(* IEC 61131-3 sources: Jacob-Formschaumtechnik-ISEL-CNC-Retrofit/twincat/PLC/src/6_Interfaces, 18 files *)

(* ---- E_AlarmId.st ---- *)
{attribute 'qualified_only'}
{attribute 'strict'}
TYPE E_AlarmId :
(
    None              := 0,
    SafetyOpen        := 100,  (* Sicherheitskreis offen / NOT-HALT *)
    DoorOpen          := 101,
    AirPressureLow    := 110,
    ExtractionFault   := 120,
    SpindleFuFault    := 200,
    SpindlePtcTrip    := 201,
    SpindleNoFeedback := 202,
    SpindleLockedSetup:= 203,
    AxisDriveFault    := 300,
    AxisFollowingErr  := 301,
    HwLimitHit        := 302,
    FieldbusLost      := 310,
    HomingLost        := 320,
    HmiLinkLost       := 330,
    ParamMismatch     := 900   (* Maschinen-ID oder Version passt nicht *)
) INT;
END_TYPE

(* ---- E_AlarmSlot.st ---- *)
{attribute 'qualified_only'}
{attribute 'strict'}
(* Meldekatalog: Slot-Nummer = Index in aCond von FB_AlarmList.
   Klassen siehe E_FaultClass. Texte und Abhilfe stehen in docs/Meldeliste.md (HMI-Thread). *)
TYPE E_AlarmSlot :
(
    SafetyOpen := 0,
    DoorOpen := 1,
    AirPressureLow := 2,
    ExtractionFault := 3,
    SpindleFuFault := 4,
    SpindlePtcTrip := 5,
    SpindleNoFeedback := 6,
    SpindleLockedSetup := 7,
    AxisDriveFault := 8,
    AxisFollowingErr := 9,
    HwLimitHit := 10,
    FieldbusLost := 11,
    HomingLost := 12,
    HmiLinkLost := 13,
    ParamMismatch := 14
) INT;
END_TYPE

(* ---- E_DriveVariant.st ---- *)
{attribute 'qualified_only'}
{attribute 'strict'}
(* Generische Achsschnittstelle. Variante A: CANopen DS402 ueber EL6751 (Interpolated Position
   unbestaetigt), Variante B: +-10 V Analog + Encoder-Klemmen (Rueckfall). *)
TYPE E_DriveVariant :
(
    CanopenDs402 := 0,
    AnalogEncoder := 1,
    Simulation := 2
) INT;
END_TYPE

(* ---- E_FaultClass.st ---- *)
{attribute 'qualified_only'}
{attribute 'strict'}
(* Fehlerreaktionsklassen, siehe docs/Architektur_Sicherheit.md *)
TYPE E_FaultClass :
(
    R0_Info     := 0,  (* nur anzeigen *)
    R1_Warning  := 1,  (* anzeigen, Betrieb laeuft weiter *)
    R2_FeedHold := 2,  (* gefuehrter Vorschubhalt, fortsetzbar *)
    R3_Abort    := 3,  (* gefuehrter Halt, Spindel aus, Programm beendet *)
    R4_DrivesOff := 4  (* Reglerfreigabe weg, Referenz verloren *)
) INT;
END_TYPE

(* ---- E_HomeState.st ---- *)
{attribute 'qualified_only'}
{attribute 'strict'}
TYPE E_HomeState :
(
    Open := 0,
    Running := 1,
    Done := 2,
    Error := 3
) INT;
END_TYPE

(* ---- E_MachState.st ---- *)
{attribute 'qualified_only'}
{attribute 'strict'}
TYPE E_MachState :
(
    Stopped     := 0,  (* Antriebe aus, kein Fehler *)
    Idle        := 1,  (* Antriebe bereit, kein Programm *)
    Execute     := 2,  (* Programm laeuft *)
    Held        := 3,  (* Vorschubhalt, Programm fortsetzbar *)
    Aborted     := 4,  (* Programm abgebrochen, Reset noetig *)
    EStop       := 5,  (* Sicherheitskreis offen *)
    Fault       := 6   (* Fehler R3/R4 aktiv, Quittierung noetig *)
) INT;
END_TYPE

(* ---- E_OpMode.st ---- *)
{attribute 'qualified_only'}
{attribute 'strict'}
TYPE E_OpMode :
(
    Hand  := 0,   (* Tippen, Handrad, Referenzieren *)
    Auto  := 1,   (* Programmbetrieb *)
    Setup := 2    (* Einrichten/Test: Spindel gesperrt, Einzelsatz moeglich *)
) INT;
END_TYPE

(* ---- ST_Alarm.st ---- *)
(* Eine Meldung aus der Meldeliste, Index = E_AlarmSlot *)
TYPE ST_Alarm :
STRUCT
    nId     : INT;
    eClass  : E_FaultClass;
    bActive : BOOL;          (* Ursache besteht *)
    bLatched: BOOL;          (* R3/R4 gespeichert, wartet auf Quittierung *)
END_STRUCT
END_TYPE

(* ---- ST_AxisMirror.st ---- *)
(* CNC-Spiegel fuer die HMI, Achsnummern der HMI: 1 = X (Quer), 2 = Y (Portal, Gantry), 3 = Z. *)
TYPE ST_AxisMirror :
STRUCT
    rActPosMach : LREAL;    (* mm, Maschinenkoordinate *)
    rActPosWork : LREAL;    (* mm, Werkstueckkoordinate *)
    bHomed      : BOOL;
END_STRUCT
END_TYPE

(* ---- ST_HmiCmd.st ---- *)
(* HMI -> SPS. Die HMI fordert nur an. Alle Verriegelungen liegen in der SPS. *)
TYPE ST_HmiCmd :
STRUCT
    nHeartbeat      : UINT;    (* Lebenszeichen, wird von der HMI hochgezaehlt *)
    eModeRequest    : E_OpMode;
    bStart          : BOOL;    (* Impuls *)
    bHold           : BOOL;    (* Impuls, Vorschubhalt *)
    bAbort          : BOOL;    (* Impuls *)
    bAck            : BOOL;    (* Impuls, Meldungen quittieren, Wiederanlauf *)
    bJogPlus        : BOOL;    (* gehalten, nur mit Heartbeat *)
    bJogMinus       : BOOL;
    nJogAxis        : USINT;   (* 1=X, 2=Y, 3=Z *)
    bJogRapid       : BOOL;
    bSpindleOn      : BOOL;    (* nur Hand *)
    bSpindleCcw     : BOOL;
    rSpindleSetRpm  : REAL;    (* 1/min *)
    bExtraction     : BOOL;
    bBlowAir        : BOOL;
    bVacuum         : BOOL;
    bHomeRequest    : BOOL;    (* Impuls *)
    bToolChangeDone : BOOL;    (* Impuls, Quittung manueller Werkzeugwechsel *)
    rJogStepMm      : REAL;    (* 0 = kontinuierlich, sonst 0.01 / 0.1 / 1 / 10 mm *)
    bHandwheelEnable: BOOL;    (* nur M1 mit Bestandsgeraet, [offen] *)
    nHandwheelAxis  : USINT;   (* 1=X, 2=Y, 3=Z *)
    nHandwheelRatio : USINT;   (* 1, 10, 100 *)
    bHomeAxis       : ARRAY[1..3] OF BOOL;   (* Impuls: einzelne Achse referenzieren *)
    bHomeAbort      : BOOL;    (* Impuls *)
    bSingleBlock    : BOOL;    (* Einzelsatz *)
    bDryRun         : BOOL;    (* Trockenlauf: Spindel gesperrt *)
    bOptStop        : BOOL;    (* optionaler Halt M1 *)
END_STRUCT
END_TYPE

(* ---- ST_HmiCncCmd.st ---- *)
(* HMI -> SPS *)
TYPE ST_HmiCncCmd :
STRUCT
    nOvrFeed       : UINT := 100;                (* % 0..120 *)
    nOvrRapid      : UINT := 100;                (* % 0..100 *)
    nOvrSpindle    : UINT := 100;                (* % 50..120 *)
    sProgramSelect : STRING(255);
    bProgramLoad   : BOOL;                       (* Impuls, nur im Stillstand *)
    aTool          : ARRAY[1..32] OF ST_Tool;    (* Schreibpuffer *)
    aWcs           : ARRAY[54..59] OF ST_Wcs;
    bTableWrite    : BOOL;                       (* Impuls: Puffer uebernehmen *)
    bWcsSetCurrent : BOOL;                       (* Impuls: aktuelle Position als Nullpunkt von nActWcs *)
    bWcsTableWrite : BOOL;                       (* Impuls: nur die Nullpunkte (G54..G59) aus aWcs uebernehmen. bTableWrite uebernimmt nur noch Werkzeuge (G-16) *)
    nSpeedLimitPct : UINT := 25;                 (* % 1..100, Inbetriebnahme-Begrenzung (Service). Wirkt nur nach unten auf Vorschub-/Eilgang-Override und Tippen. Anheben nur im Stillstand. *)
END_STRUCT
END_TYPE

(* ---- ST_HmiCncSts.st ---- *)
(* SPS -> HMI *)
TYPE ST_HmiCncSts :
STRUCT
    aAxis         : ARRAY[1..3] OF ST_AxisMirror;
    rGantryDiffMm : LREAL;                       (* Y1 minus Y2 *)
    nOvrFeed      : UINT;                        (* % *)
    nOvrRapid     : UINT;
    nOvrSpindle   : UINT;
    sProgramName  : STRING(80);
    nActBlock     : UDINT;
    nTotalBlocks  : UDINT;
    sBlockText    : ARRAY[0..6] OF STRING(80);   (* Index 3 = aktueller Satz *)
    rRestMm       : LREAL;
    rFeedAct      : LREAL;                       (* mm/min *)
    nActTool      : UINT;
    nActWcs       : UINT := 54;                  (* 54..59 *)
    aTool         : ARRAY[1..32] OF ST_Tool;
    aWcs          : ARRAY[54..59] OF ST_Wcs;
    bProgramLoaded: BOOL;
    bTableWriteOk : BOOL;                        (* Rueckmeldung letzter Schreibvorgang *)
    bTableWriteRejected : BOOL;                  (* abgelehnt, z. B. Programm laeuft *)
    nSpeedLimitActivePct : UINT := 25;           (* wirksame Inbetriebnahme-Begrenzung in %, nOvrFeed/nOvrRapid sind bereits damit begrenzt *)
END_STRUCT
END_TYPE

(* ---- ST_HmiJournal.st ---- *)
(* Meldejournal fuer die HMI (Befund 21, LH-2.9.2). Ringpuffer der letzten 100 kommenden Meldungen.
   nHead zeigt auf den naechsten freien Platz, der juengste Eintrag steht bei (nHead + 99) MOD 100.
   nSeq zaehlt jeden neuen Eintrag hoch, die HMI liest nur bei Aenderung. *)
TYPE ST_HmiJournal :
STRUCT
    aEntry   : ARRAY[0..99] OF ST_JournalEntry;
    nHead    : UINT;
    nEntries : UINT;
    nSeq     : UDINT;
END_STRUCT
END_TYPE

(* ---- ST_HmiSts.st ---- *)
(* SPS -> HMI. CNC-Werte (Achspositionen, Overrides, Werkzeug-/Nullpunkttabelle) liefert der
   CNC-Spiegel GVL_HmiCnc (ST_HmiCncSts), solange TF5310 nicht verfuegbar ist. *)
TYPE ST_HmiSts :
STRUCT
    eMode           : E_OpMode;
    eState          : E_MachState;
    bSafetyOk       : BOOL;
    bDrivesEnabled  : BOOL;
    bAllHomed       : BOOL;
    bHmiLinkOk      : BOOL;    (* Heartbeat der HMI wird ueberwacht *)
    bSpindleRunning : BOOL;
    rSpindleActRpm  : REAL;
    bExtractionOn   : BOOL;
    bBlowAirOn      : BOOL;
    bVacuumOn       : BOOL;
    bToolChangeReq  : BOOL;    (* Aufforderung am Panel *)
    nToolChangeNo   : UINT;
    nTopAlarmId     : INT;     (* hoechste aktive Meldung, 0 = keine *)
    eTopAlarmClass  : E_FaultClass;
    nActiveAlarms   : UINT;
    nMachineId      : UINT;    (* aus Maschinenparametern, z. B. 1 fuer M1 *)
    sSwVersion      : STRING(15);
    dwOperatingSec  : UDINT;   (* Betriebssekunden, fuer Wartungsanzeige *)
    dwSpindleSec    : UDINT;
    bHandwheelActive: BOOL;
    eHomeState      : ARRAY[1..3] OF E_HomeState;
    nHomeStep       : USINT;
    aAlarms         : ARRAY[0..14] OF ST_Alarm;    (* Index = E_AlarmSlot *)
    aDrive          : ARRAY[1..4] OF ST_AxisDrive; (* Diagnose, 1=Y1 2=Y2 3=X 4=Z [Annahme] *)
    bFieldbusOk     : BOOL;
    bFuFault        : BOOL;    (* Rohsignal *)
    bPtcTrip        : BOOL;    (* Rohsignal *)
    bSimulationActive : BOOL;  (* Simulationsabbild der Antriebe aktiv, nie auf einer realen Maschine *)
    bModeChangeBlocked: BOOL;  (* Betriebsartenwunsch abgelehnt *)
    nHeartbeatEcho  : UINT;    (* Rueckspiegel stCmd.nHeartbeat, Befund 16 *)
    bLimitFreeRun   : BOOL;    (* Endschalter angefahren, Freifahren in Hand im Schleichgang moeglich, Befund 15 *)
    bToolChangeDoorRelease : BOOL;  (* Werkzeugwechsel: Spindel steht, Tuer darf geoeffnet werden *)
END_STRUCT
END_TYPE

(* ---- ST_JournalEntry.st ---- *)
(* Eintrag im Meldejournal (Befund 21). Zeitstempel in UTC. *)
TYPE ST_JournalEntry :
STRUCT
    nId    : INT;      (* Meldungs-ID aus GVL_AlarmCatalog *)
    nClass : INT;      (* 0..4 = R0..R4 *)
    dtTime : DT;       (* Kommt-Zeitpunkt, UTC *)
END_STRUCT
END_TYPE

(* ---- ST_MachineParams.st ---- *)
(* Maschinenparameter. Je Maschine eine Datei in config/, geladen beim Start.
   Werte in config/M1.json mit [Annahme] gekennzeichnet, solange nicht bestaetigt. *)
TYPE ST_MachineParams :
STRUCT
    nMachineId        : UINT;
    sSwVersionExpected: STRING(15);
    eDriveVariant     : E_DriveVariant;    (* muss zur Build-Konfiguration passen (Befund 20) *)
    nNumAxes          : USINT;             (* Antriebe ohne Spindel: Y1, Y2, X, Z = 4 *)
    nNumCncAxes       : USINT;             (* CNC-/HMI-Achsen X, Y, Z = 3 (Y als Gantry) *)
    rSpindleMaxRpm    : REAL;              (* 16600 fuer VKH63/26-90T *)
    rSpindleMinRpm    : REAL;
    rSpindleVoltMax   : REAL;              (* 10.0 V entspricht rSpindleMaxRpm *)
    tSpindleRunUp     : TIME;              (* Wartezeit nach Start bis Drehzahl erreicht *)
    tSpindleStandstill: TIME;              (* Auslaufzeit bis Stillstand gemeldet *)
    tHmiTimeout       : TIME;              (* Heartbeat-Ausfall -> Tippen stoppt *)
    tFeedbackTimeout  : TIME;              (* Rueckmeldung Ventil/Spindel *)
    bAirMonitoring    : BOOL;
    bHasToolChanger   : BOOL;
END_STRUCT
END_TYPE

(* ---- ST_Tool.st ---- *)
TYPE ST_Tool :
STRUCT
    nNo     : UINT;
    sName   : STRING(31);
    rLength : LREAL;        (* mm *)
    rRadius : LREAL;        (* mm *)
END_STRUCT
END_TYPE

(* ---- ST_Wcs.st ---- *)
TYPE ST_Wcs :
STRUCT
    rX : LREAL;             (* mm, Nullpunktverschiebung *)
    rY : LREAL;
    rZ : LREAL;
END_STRUCT
END_TYPE
